// TIA Portal V18 export
FUNCTION_BLOCK "EmptyPhase"   // FB101, SCL
{ S7_Optimized_Access := 'TRUE' }
VERSION : 0.1
// stored: AutoNumber true, IsIECCheckEnabled false, IsRetainMemResEnabled false, MemoryReserve 100, SetENOAutomatically false, UDAEnableTagReadback false
   VAR_INPUT
      SP01 { ExternalAccessible := 'False'; ExternalVisible := 'False'; ExternalWritable := 'False'} : Real;
      SP02 { ExternalAccessible := 'False'; ExternalVisible := 'False'; ExternalWritable := 'False'} : Real;
      SP03 { ExternalAccessible := 'False'; ExternalVisible := 'False'; ExternalWritable := 'False'} : Real;
      SP04 { ExternalAccessible := 'False'; ExternalVisible := 'False'; ExternalWritable := 'False'} : Real;
      SP05 { ExternalAccessible := 'False'; ExternalVisible := 'False'; ExternalWritable := 'False'} : Real;
      InterfaceIn { ExternalAccessible := 'False'; ExternalVisible := 'False'; ExternalWritable := 'False'} : DWord;
   END_VAR
   VAR_OUTPUT
      IDLE { ExternalAccessible := 'False'; ExternalVisible := 'False'; ExternalWritable := 'False'} : Bool;
      HELD { ExternalAccessible := 'False'; ExternalVisible := 'False'; ExternalWritable := 'False'} : Bool;
      START { ExternalAccessible := 'False'; ExternalVisible := 'False'; ExternalWritable := 'False'} : Bool;
      STOP { ExternalAccessible := 'False'; ExternalVisible := 'False'; ExternalWritable := 'False'} : Bool;
      ABORT { ExternalAccessible := 'False'; ExternalVisible := 'False'; ExternalWritable := 'False'} : Bool;
      PAUSE { ExternalAccessible := 'False'; ExternalVisible := 'False'; ExternalWritable := 'False'} : Bool;
      PAUSING { ExternalAccessible := 'False'; ExternalVisible := 'False'; ExternalWritable := 'False'} : Bool;
      STARTING { ExternalAccessible := 'False'; ExternalVisible := 'False'; ExternalWritable := 'False'} : Bool;
      STOPPING { ExternalAccessible := 'False'; ExternalVisible := 'False'; ExternalWritable := 'False'} : Bool;
      ABORTING { ExternalAccessible := 'False'; ExternalVisible := 'False'; ExternalWritable := 'False'} : Bool;
      COMPLETED { ExternalAccessible := 'False'; ExternalVisible := 'False'; ExternalWritable := 'False'} : Bool;
      InterfaceOut { ExternalAccessible := 'False'; ExternalVisible := 'False'; ExternalWritable := 'False'} : DWord;
   END_VAR
   VAR_IN_OUT
      InterfaceInOut { ExternalAccessible := 'False'; ExternalVisible := 'False'; ExternalWritable := 'False'} : DWord;
   END_VAR
   VAR
      "timer" : "fbTimer";
      "step" { ExternalAccessible := 'False'; ExternalVisible := 'False'; ExternalWritable := 'False'} : Int;
      step_prev { ExternalAccessible := 'False'; ExternalVisible := 'False'; ExternalWritable := 'False'} : Int;
      count : USInt;
      ALARM_BLOCK { ExternalAccessible := 'False'; ExternalVisible := 'False'; ExternalWritable := 'False'} : "AlarmBlock";
      AlarmBlock { ExternalAccessible := 'False'; ExternalVisible := 'False'; ExternalWritable := 'False'} : Program_Alarm;
      Message_1 { ExternalAccessible := 'False'; ExternalVisible := 'False'; ExternalWritable := 'False'} : Program_Alarm;
      Message_2 { ExternalAccessible := 'False'; ExternalVisible := 'False'; ExternalWritable := 'False'} : Program_Alarm;
      Message_3 { ExternalAccessible := 'False'; ExternalVisible := 'False'; ExternalWritable := 'False'} : Program_Alarm;
      Message_4 { ExternalAccessible := 'False'; ExternalVisible := 'False'; ExternalWritable := 'False'} : Program_Alarm;
      Message_5 { ExternalAccessible := 'False'; ExternalVisible := 'False'; ExternalWritable := 'False'} : Program_Alarm;
      OpRequest_1 : "fbOpMsg";
      OpRequest_2 : "fbOpMsg";
      OpRequest_3 : "fbOpMsg";
      OpRequest_4 : "fbOpMsg";
      OpRequest_5 : "fbOpMsg";
      TRANSFER : "fbTransfer";
      TRANSFER_READY { ExternalAccessible := 'False'; ExternalVisible := 'False'; ExternalWritable := 'False'} : Bool;
   END_VAR
   // ALARM_BLOCK.TEXTLIST_ID := 519;
   // ALARM_BLOCK.INDEX := 0;
BEGIN
   REGION COMMANDS
       #STOP := #InterfaceIn.%X12;
       #IDLE := #InterfaceIn.%X11;
       #HELD := #InterfaceIn.%X10;
       #START := #InterfaceIn.%X16;
       #ABORT := #InterfaceIn.%X14;
       #PAUSE := #InterfaceIn.%X13;
       #ABORTING := #InterfaceIn.%X21;
       #STARTING := #InterfaceIn.%X20;
       #STOPPING := #InterfaceIn.%X19;
   END_REGION
   REGION FUNCTION
       IF #START OR #PAUSE THEN

           //======================================================================================================================
           IF #STARTING THEN
               #step := 10;
               #count := 0;

               #Message_1.SIG := false;
               #Message_2.SIG := false;
               #Message_3.SIG := false;
               #Message_4.SIG := false;
               #Message_5.SIG := false;

               #TRANSFER_READY := false;

           ELSIF #START THEN
               ;
           END_IF;

           //======================================================================================================================

           CASE #step OF

               10:  // =============================================================================================================
                   REGION S10 -   
                       //Action

                       //Next
                       IF false THEN
                           IF NOT #PAUSE THEN
                               #step += 10;
                           END_IF;
                       END_IF;
                   END_REGION

               20:  // =============================================================================================================
                   REGION S20 -   
                       //Action

                       //Next
                       #COMPLETED := true;
                   END_REGION
           END_CASE;

       ELSIF #STOP THEN
           IF #STOPPING THEN
               ;
           END_IF;
           #TRANSFER_READY := false;
       ELSIF #ABORT THEN
           #COMPLETED := false;
       END_IF;

   END_REGION

   REGION MESSAGES
       #Message_1();
       #Message_2();
       #Message_3();
       #Message_4();
       #Message_5();
   END_REGION

   REGION OPERATOR REQUEST
       #OpRequest_1(MESSAGE := #START AND #step = -1,
                    "TYPE" := 0);

       #OpRequest_2(MESSAGE := #START AND #step = -1,
                    "TYPE" := 0);

       #OpRequest_3(MESSAGE := #START AND #step = -1,
                    "TYPE" := 0);

       #OpRequest_4(MESSAGE := #START AND #step = -1,
                    "TYPE" := 0);

       #OpRequest_5(MESSAGE := #START AND #step = -1,
                    "TYPE" := 0);

   END_REGION

   REGION TRANSFER
       #TRANSFER(BIT_READY:=#TRANSFER_READY AND NOT #HELD);

       IF #TRANSFER.ACTIVE THEN
           ;
       ELSIF #TRANSFER.READY OR #TRANSFER.HELD OR #TRANSFER.COMPLETED THEN
           ;
       END_IF;
   END_REGION

   REGION TIMER
       IF NOT #START OR #START AND #step <> #step_prev THEN
           #timer.Start := false;
       END_IF;

       #timer();
   END_REGION

   REGION STATUS
       IF FALSE THEN
           #InterfaceOut.%X24 := true;
       ELSE
           #InterfaceOut.%X24 := false;
       END_IF;

       #InterfaceOut.%X22 := #COMPLETED;
       #InterfaceOut.%X23 := #STOP OR #IDLE;
       #InterfaceOut.%X25 := #OpRequest_1.Interface = -1 OR #OpRequest_2.Interface = -1 OR #OpRequest_3.Interface = -1 OR #OpRequest_4.Interface = -1 OR #OpRequest_5.Interface = -1;

       #AlarmBlock(SIG := #HELD,
                   SD_1 := #ALARM_BLOCK.TEXTLIST_ID,
                   SD_2 := #ALARM_BLOCK.INDEX);

       IF NOT #IDLE THEN
           #InterfaceInOut.%X10 := true;
       END_IF;

       IF #HELD THEN
           #InterfaceInOut.%X11 := true;
       END_IF;

       IF #START THEN
           #InterfaceInOut.%X12 := true;
       END_IF;

       IF #STOP THEN
           #InterfaceInOut.%X13 := true;
       END_IF;

       IF #ABORT THEN
           #InterfaceInOut.%X14 := true;
       END_IF;

       IF #PAUSE THEN
           #InterfaceInOut.%X15 := true;
       END_IF;

       IF #COMPLETED THEN
           #InterfaceInOut.%X16 := true;
       END_IF;

       #step_prev := #step;
   END_REGION
END_FUNCTION_BLOCK
